// TwinCAT 3 PLC project LibraryDocumentationSample
// Title: LibraryDocumentationSample
// Company: Beckhoff Automation GmbH & Co. KG
// ProjectVersion: 1.0.0.0
// Description: This library contains various function blocks ...
// ProgramVersion: 3.1.4026.25
// project tree:
//   LibPOUs/A_Samples/ FB_DocuSample_FunctionBlock.TcPOU, FB_DocuSample_SyntaxReminder.TcPOU
//   LibPOUs/B_DocuElements/Code block/ FB_Libdoc_CodeBlock.TcPOU
//   LibPOUs/B_DocuElements/Hyperlinks/ FB_Libdoc_LinkToAnotherObject.TcPOU, FB_Libdoc_AnonymousHyperlinks.TcPOU, FB_Libdoc_Citation.TcPOU, FB_Libdoc_ExternalHyperlinks.TcPOU, FB_Libdoc_IndirectHyperlinks.TcPOU, FB_Libdoc_InlineHyperlinks.TcPOU, FB_Libdoc_InternalHyperlinks.TcPOU
//   LibPOUs/B_DocuElements/Internal Comments/ FB_Libdoc_InternalComments.TcPOU
//   LibPOUs/B_DocuElements/Font style/ FB_Libdoc_FontStyle.TcPOU
//   LibPOUs/B_DocuElements/Hyperlinks/Footnotes/ FB_Libdoc_AutomaticallyNumberedFootnotes.TcPOU, FB_Libdoc_AutomaticallySymbolFootnotes.TcPOU, FB_Libdoc_ManuallyAndAutomaticallyNumberedFootnotes.TcPOU, FB_Libdoc_ManuallyNumberedFootnotes.TcPOU, FB_Libdoc_NamedAutomaticallyNumberedFootnotes.TcPOU
//   LibPOUs/B_DocuElements/Images/ FB_Libdoc_Images.TcPOU
//   LibPOUs/B_DocuElements/Lists/ FB_Libdoc_DefinitionList.TcPOU, FB_Libdoc_FieldList.TcPOU, FB_Libdoc_OrderedNumberedEnumerationList.TcPOU, FB_Libdoc_UnorderedEnumerationList.TcPOU
//   LibPOUs/B_DocuElements/Note elements/ FB_Libdoc_SpecificNotes.TcPOU, FB_Libdoc_GenericNotes.TcPOU
//   LibPOUs/B_DocuElements/Comment structure/ FB_Libdoc_Sections.TcPOU, FB_Libdoc_Transitions.TcPOU
//   LibPOUs/B_DocuElements/Substitution/ FB_Libdoc_Substitution_ReplacementText.TcPOU, FB_Libdoc_Substitution_Images.TcPOU
//   LibPOUs/B_DocuElements/Tables/ FB_Libdoc_CSVTable.TcPOU, FB_Libdoc_GridTable.TcPOU, FB_Libdoc_ListTable.TcPOU, FB_Libdoc_SimpleTables.TcPOU
//   LibPOUs/B_DocuElements/Text blocks/ FB_Libdoc_LineBlock.TcPOU, FB_Libdoc_Paragraph.TcPOU, FB_Libdoc_BlockQuote.TcPOU

// ---- LibPOUs/A_Samples/FB_DocuSample_FunctionBlock.TcPOU
(* 
:Description: This function block represents <...> and can be used for <...> ...
:Instructions for use: How to use this FB ...

Version history:

+-------------+------------+----------------+----------+------------------------------------------+
|Date         | Version    | created under  | Author   | Remark                                   |
+=============+============+================+==========+==========================================+
|2017-07-04   | 1.0.0.0    | V3.1.4022.0    | S.H.     | Performance optimization                 |
+-------------+------------+----------------+----------+------------------------------------------+
|2019-01-11   | 1.1.0.0    | V3.1.4022.27   | K.F.     | Bug fix: Output calculation corrected    |
+-------------+------------+----------------+----------+------------------------------------------+
*)

FUNCTION_BLOCK FB_DocuSample_FunctionBlock
VAR_INPUT
    nVarInA : INT;       //First input variable
    nVarInB : INT := 5;  //Second input variable
END_VAR
VAR_OUTPUT
    nVarOut : INT;       //Output variable
END_VAR

END_FUNCTION_BLOCK

// ---- LibPOUs/A_Samples/FB_DocuSample_SyntaxReminder.TcPOU
(*
=================================================
The reStructuredText Cheat Sheet: Syntax Reminder
=================================================
:Info: See <https://infosys.beckhoff.de/.
:Author: Beckhoff <support@beckhoff.com>
:Date: 2017-12-14

.. NOTE:: This syntax reminder is based on the docutils documentation

Section Structure
=================

A reStructuredText comment is made up of body elements, and may be
structured into sections. Section titles are underlined or overlined and underlined.
Sections contain body elements and/or subsections.

Paragraphs are flush-left and separated by blank lines.

Body Elements
=============
Grid table:

+--------------------------------+-------------------------------------+
|Block quotes consist of         |Literal block, preceded by "::"::    |
|indented body elements:         |                                     |
|                                |    If (a=TRUE) Then                 |
|    Block quotes are indented.  |      b=3                            |
|                                |                                     |
+--------------------------------+-------------------------------------+
|| Line blocks preserve line breaks and indents.                       |
||    Useful for adornment-free lists;                                 |
||    long lines can be wrapped                                        |
|     with continuation lines.                                         |
+----------------------------------------------------------------------+

Simple table:

================  ========================================================
List Type         Examples
================  ========================================================
Bullet list       - This is a bullet list
                  - Items begin with "-", "+", or "*"
Enumerated list   1. This is an enumerated list.
                  2. Items use any variation of "1.", "A)", and "(i)"
                  #. Item can also be auto-enumerated
Definition list   Term is flush-left : optional classifier
                      Definition is indented, no blank line between
                      continue
Field list        :Field name: field body
================  ========================================================

Inline Markup
=============
*emphasis*, **strong emphasis**, ``inline literal text``

| Standalone hyperlink: http://beckhoff.de
| Named reference: Beckhoff_
| Anonymous reference: `Anonymous reference`__
| Footnote reference: [1]_
| Citation reference: [CIT2002]_
| Substitution: |substitution|
| Inline internal target: `Inline internal target`_

Explicit Markup
================

================  ========================================================
Explicit Markup       Examples (visible in the source code)
================  ========================================================
Footnote          .. [1] Manually numbered or [#] auto-numbered
                        (even [#label]) or [*] auto-symbol
Citation          .. [CIT2002] This is a citation.
Hyperlink Target  .. _Beckhoff: http://beckhoff.de
                  .. _indirect target: Beckhoff_
                  .. _internal target:
Anonymous Target  __ http://beckhoff.de
Directive ("::")  .. image::, .. code::
Substitution Def  .. |substitution| replace:: This is a substitution
Comment           .. This text will not be shown
================  ========================================================

Directives
===========

================  ========================================================
Directive Name    Description
================  ========================================================
attention         Specific admonition ("caution", "danger",
                  "error", "hint", "important", "note", "tip", "warning")
admonition        Generic titled admonition
image             .. image:: C:\Tc3LibDocImages\BeckhoffLogo.png
                     :width: 40
code              .. code::

                     if(a=true) then b=3;
list-table        Create a table from a uniform two-level bullet list
csv-table         Create a table from CSV data
================  ========================================================*)

FUNCTION_BLOCK FB_DocuSample_SyntaxReminder
VAR_INPUT
    nVarInA : INT;       //First input variable
    nVarInB : INT := 5;  //Second input variable
END_VAR
VAR_OUTPUT
    nVarOut : INT;       //Output variable
END_VAR

END_FUNCTION_BLOCK

// ---- LibPOUs/B_DocuElements/Code block/FB_Libdoc_CodeBlock.TcPOU
(*

**Code block with color-coded syntax**

.. code:: 
    
    // Attempts to return the value of a boolean property.
   
    FUNCTION GetBooleanProperty : BOOL
    VAR_INPUT
        sKey: STRING;
    END_VAR

    // This structure defines a special profile.

    TYPE ST_Profile :
    STRUCT
        nId     : INT := -1;
        sBuffer : STRING(255) := 'Hello';
    END_STRUCT
    END_TYPE

**Code block with line numbering**

.. code:: 
   :number-lines: 1
    
    // Attempts to return the value of a boolean property.
   
    FUNCTION GetBooleanProperty : BOOL
    VAR_INPUT
        sKey: STRING;
    END_VAR

    // This structure defines a special profile.

    TYPE ST_Profile :
    STRUCT
        nId     : INT := -1;
        sBuffer : STRING(255) := 'Hello';
    END_STRUCT
    END_TYPE

*)

FUNCTION_BLOCK FB_Libdoc_CodeBlock
VAR_INPUT
    nVarA : INT;
    nVarB : INT;
END_VAR
VAR_OUTPUT
    nSum : INT;
END_VAR
VAR
END_VAR

END_FUNCTION_BLOCK

// ---- LibPOUs/B_DocuElements/Hyperlinks/FB_Libdoc_LinkToAnotherObject.TcPOU
(*
| It is also possible to create a reference to the documentation of another object which is also part of this library.
| For example, by clicking on this link :ref:`FB_Libdoc_InlineHyperlinks`, the documentation of this FB will be shown.
| Or you can also create a link to :ref:`FB_Libdoc_CodeBlock` which is part of another folder.

*)

FUNCTION_BLOCK FB_Libdoc_LinkToAnotherObject
VAR_INPUT
    nVarA : INT;
    nVarB : INT;
END_VAR
VAR_OUTPUT
    nSum : INT;
END_VAR
VAR
END_VAR

END_FUNCTION_BLOCK

// ---- LibPOUs/B_DocuElements/Internal Comments/FB_Libdoc_InternalComments.TcPOU
(*
This is the first paragraph.

.. Comments begin with two dots and one space. Anything can
   follow, except for the syntax of footnotes/citations,
   hyperlink targets, directives, or substitution definitions.

Since comments are not shown, this paragraph follows the previous paragraph directly.
*)

FUNCTION_BLOCK FB_Libdoc_InternalComments
VAR_INPUT
    nVarA : INT;
    nVarB : INT;
END_VAR
VAR_OUTPUT
    nSum : INT;
END_VAR
VAR
END_VAR

END_FUNCTION_BLOCK

// ---- LibPOUs/B_DocuElements/Font style/FB_Libdoc_FontStyle.TcPOU
(*
This is *emphasized text*.

This is **strong text**.

This text is an example of ``inline literals``.
*)

FUNCTION_BLOCK FB_Libdoc_FontStyle
VAR_INPUT
    nVarA : INT;
    nVarB : INT;
END_VAR
VAR_OUTPUT
    nSum : INT;
END_VAR
VAR
END_VAR

END_FUNCTION_BLOCK

// ---- LibPOUs/B_DocuElements/Hyperlinks/FB_Libdoc_AnonymousHyperlinks.TcPOU
(*
See the `Beckhoff Online Information System`__ or the `Beckhoff home page`__.

.. __: http://infosys.beckhoff.de/

.. __: http://beckhoff.de/
*)

FUNCTION_BLOCK FB_Libdoc_AnonymousHyperlinks
VAR_INPUT
    nVarA : INT;
    nVarB : INT;
END_VAR
VAR_OUTPUT
    nSum : INT;
END_VAR
VAR
END_VAR

END_FUNCTION_BLOCK

// ---- LibPOUs/B_DocuElements/Hyperlinks/FB_Libdoc_Citation.TcPOU
(*
Citation references, like [CIT2002]_. Note that citations may get rearranged, e.g., to the bottom of the "page". 

| Some sample text to get some text in between.
| Some sample text to get some text in between.
| Some sample text to get some text in between.
| Some sample text to get some text in between.
| Some sample text to get some text in between.
| Some sample text to get some text in between.

.. [CIT2002] This is the citation.  It's just like a footnote,
   except the label is textual. 

Given a citation like [this]_, one can also refer to it like this_. 

| Some sample text to get some text in between.
| Some sample text to get some text in between.
| Some sample text to get some text in between.
| Some sample text to get some text in between.
| Some sample text to get some text in between.
| Some sample text to get some text in between.

.. [this] here.

| Some sample text to get some text in between.
| Some sample text to get some text in between.
| Some sample text to get some text in between.
| Some sample text to get some text in between.
| Some sample text to get some text in between.
| Some sample text to get some text in between.

*)

FUNCTION_BLOCK FB_Libdoc_Citation
VAR_INPUT
    nVarA : INT;
    nVarB : INT;
END_VAR
VAR_OUTPUT
    nSum : INT;
END_VAR
VAR
END_VAR

END_FUNCTION_BLOCK

// ---- LibPOUs/B_DocuElements/Hyperlinks/FB_Libdoc_ExternalHyperlinks.TcPOU
(*
See the Beckhoff homepage_ for more information.

Please contact the `Beckhoff Support`_ for technical assistance.

.. _homepage: http://www.beckhoff.de
.. _Beckhoff Support: support@beckhoff.com

For more information see the `PLC Lib Tc2_System`_ and `PLC Lib Tc2_Standard`_.

.. _PLC Lib Tc2_System: https://download.beckhoff.com/download/document/automation/twincat3/TwinCAT_3_PLC_Lib_Tc2_System_EN.pdf
.. _PLC Lib Tc2_Standard: https://download.beckhoff.com/download/document/automation/twincat3/TwinCAT_3_PLC_Lib__Tc2_Standard_EN.pdf

External hyperlinks, like `Beckhoff <http://www.beckhoff.de/>`_.


**Standalone hyperlinks**

See http://www.beckhoff.de for info.

Contact support@beckhoff.com


**Embedded URIs and aliases**

See the `Beckhoff homepage <http://www.beckhoff.de>`_ for info.

This `link <Beckhoff homepage_>`_ is an alias to the link above.


See the `Beckhoff homepage`_ for info.

This link_ is an alias to the link above.

.. _Beckhoff homepage: http://www.beckhoff.de
.. _link: `Beckhoff homepage`_

*)

FUNCTION_BLOCK FB_Libdoc_ExternalHyperlinks
VAR_INPUT
    nVarA : INT;
    nVarB : INT;
END_VAR
VAR_OUTPUT
    nSum : INT;
END_VAR
VAR
END_VAR

END_FUNCTION_BLOCK

// ---- LibPOUs/B_DocuElements/Hyperlinks/FB_Libdoc_IndirectHyperlinks.TcPOU
(*

**Indirect references to an internal reference target**

This hyperlink points to target one_ and indirect to target three.

.. _one: two_
.. _two: three_
.. _three:

The hyperlink targets above point to this paragraph.

**Indirect references to an external reference target**

The `Beckhoff Information System`_ is a reference source for Beckhoff_ products

.. _Beckhoff: `Beckhoff Information System`_

.. _Beckhoff Information System: https://infosys.beckhoff.de/
*)

FUNCTION_BLOCK FB_Libdoc_IndirectHyperlinks
VAR_INPUT
    nVarA : INT;
    nVarB : INT;
END_VAR
VAR_OUTPUT
    nSum : INT;
END_VAR
VAR
END_VAR

END_FUNCTION_BLOCK

// ---- LibPOUs/B_DocuElements/Hyperlinks/FB_Libdoc_InlineHyperlinks.TcPOU
(*
| This function block is based on a _`statemachine` concept which is described in the following.
| The statemachine is based on several states.
| The proceeding always begins in the first state.
| If the last state is left, the execution restarts in the first state.
| There are so many more information necessary to describe the statemachine concept in detail.
| But as this is just a sample text to show the inline hyperlinks, we want to leave out the details.
| A rough description should be enough for the sample demonstration.
| 
| Some sample text to get some text in between.
| Some sample text to get some text in between.
| Some sample text to get some text in between.
| Some sample text to get some text in between.
| Some sample text to get some text in between.
| Some sample text to get some text in between.
| 
| Furthermore, the function block is based on another concept. This is called XY.
| It is always necessary to respect the demands of this concept.
| Especially, as it is deeply interwoven with the statemachine concept.
| Therefore, you definitely need to understand the statemachine concept first.
| Afterwards, you might understand the XY concept.
| For more information about this, see the description of the `statemachine`_.
| By clicking on this link, the Library Manager will jump to the beginning of the first paragraph where the statemachine concept is described.. 

*)

FUNCTION_BLOCK FB_Libdoc_InlineHyperlinks
VAR_INPUT
    nVarA : INT;
    nVarB : INT;
END_VAR
VAR_OUTPUT
    nSum : INT;
END_VAR
VAR
END_VAR

END_FUNCTION_BLOCK

// ---- LibPOUs/B_DocuElements/Hyperlinks/FB_Libdoc_InternalHyperlinks.TcPOU
(*

**Simple internal hyperlink target**

Clicking on this internal hyperlink will take us to the target_
below.

.. _target:

**Nesting of internal hyperlink targets**

Clicking on this internal hyperlink will take us to the `third item`_ of the bullet list.

* First list item
* Second list item

  .. _third item:

* Third list item, with hyperlink target.

**Concatentation of internal hyperlink targets**

Clicking on this internal hyperlink will take us to target1_
and clicking on this internal hyperlink will take us to target2_.
Both targets point the the same paragraph.

.. _target1:
.. _target2:

The targets "target1" and "target2" are synonyms; they both
point to this paragraph.
*)

FUNCTION_BLOCK FB_Libdoc_InternalHyperlinks
VAR_INPUT
    nVarA : INT;
    nVarB : INT;
END_VAR
VAR_OUTPUT
    nSum : INT;
END_VAR
VAR
END_VAR

END_FUNCTION_BLOCK

// ---- LibPOUs/B_DocuElements/Hyperlinks/Footnotes/FB_Libdoc_AutomaticallyNumberedFootnotes.TcPOU
(*

**Autonumbered footnotes**

Autonumbered footnotes are possible, like using [#]_ and [#]_. 

--------

.. [#] This is the first one. 

.. [#] This is the second one. 
*)

FUNCTION_BLOCK FB_Libdoc_AutomaticallyNumberedFootnotes
VAR_INPUT
    nVarA : INT;
    nVarB : INT;
END_VAR
VAR_OUTPUT
    nSum : INT;
END_VAR
VAR
END_VAR

END_FUNCTION_BLOCK

// ---- LibPOUs/B_DocuElements/Hyperlinks/Footnotes/FB_Libdoc_AutomaticallySymbolFootnotes.TcPOU
(*

Here is a symbolic 
footnote reference: [*]_ footnote reference: [*]_
footnote reference: [*]_ footnote reference: [*]_
footnote reference: [*]_ footnote reference: [*]_
footnote reference: [*]_ footnote reference: [*]_
footnote reference: [*]_ footnote reference: [*]_
footnote reference: [*]_

.. [*] This is the first footnote.
.. [*] This is the second footnote.
.. [*] This is the third footnote.
.. [*] This is the fourth footnote.
.. [*] This is the fifth footnote.
.. [*] This is the sixth footnote.
.. [*] This is the seventh footnote.
.. [*] This is the eighth footnote.
.. [*] This is the ninth footnote.
.. [*] This is the tenth footnote.
.. [*] This is the eleventh footnote.
*)

FUNCTION_BLOCK FB_Libdoc_AutomaticallySymbolFootnotes
VAR_INPUT
    nVarA : INT;
    nVarB : INT;
END_VAR
VAR_OUTPUT
    nSum : INT;
END_VAR
VAR
END_VAR

END_FUNCTION_BLOCK

// ---- LibPOUs/B_DocuElements/Hyperlinks/Footnotes/FB_Libdoc_ManuallyAndAutomaticallyNumberedFootnotes.TcPOU
(*

[2]_ will be "2" (manually numbered footnote),

[3]_ will be "3" (another manually numbered footnote),

[#]_ will be "4" (anonymous auto-numbered footnote), and

[#label]_ will be "1" (labeled auto-numbered).

--------

.. [2] This footnote is labeled manually, so its number is fixed.

.. [3] This footnote is also labeled manually, so its number is also fixed.

.. [#label] This autonumber-labeled footnote will be labeled "1".
   It is the first auto-numbered footnote and no other footnote
   with label "1" exists.  The order of the footnotes is used to
   determine numbering, not the order of the footnote references!

.. [#] This footnote will be labeled "4".  It is the second
   auto-numbered footnote, but footnote labels "1", "2", "3" are already used. 
*)

FUNCTION_BLOCK FB_Libdoc_ManuallyAndAutomaticallyNumberedFootnotes
VAR_INPUT
    nVarA : INT;
    nVarB : INT;
END_VAR
VAR_OUTPUT
    nSum : INT;
END_VAR
VAR
END_VAR

END_FUNCTION_BLOCK

// ---- LibPOUs/B_DocuElements/Hyperlinks/Footnotes/FB_Libdoc_ManuallyNumberedFootnotes.TcPOU
(*

**Numerical footnote**

Footnote references, like [5]_. Note that footnotes may get rearranged, e.g., to the bottom of the "page".

--------

.. [5] A numerical footnote. Note there's no colon after the ``]``.
*)

FUNCTION_BLOCK FB_Libdoc_ManuallyNumberedFootnotes
VAR_INPUT
    nVarA : INT;
    nVarB : INT;
END_VAR
VAR_OUTPUT
    nSum : INT;
END_VAR
VAR
END_VAR

END_FUNCTION_BLOCK

// ---- LibPOUs/B_DocuElements/Hyperlinks/Footnotes/FB_Libdoc_NamedAutomaticallyNumberedFootnotes.TcPOU
(*

**Autonumbered labeled footnotes**

They may be assigned 'autonumber labels' - for instance, [#first]_ and [#second]_. 

--------

.. [#first] a.k.a. first_ 

.. [#second] a.k.a. second_
*)

FUNCTION_BLOCK FB_Libdoc_NamedAutomaticallyNumberedFootnotes
VAR_INPUT
    nVarA : INT;
    nVarB : INT;
END_VAR
VAR_OUTPUT
    nSum : INT;
END_VAR
VAR
END_VAR

END_FUNCTION_BLOCK

// ---- LibPOUs/B_DocuElements/Images/FB_Libdoc_Images.TcPOU
(*

**Absolute or relative file path as directive argument**

Absolute path

.. image:: C:\Tc3LibDocImages\tulpis.jpg
   :width: 70px

Relative path

.. image:: ../../LibPics/penguins.jpg
   :width: 70px

**Left aligned image**

.. image:: ../../LibPics/desert.jpg
   :width: 20%

Description of the function block. Description of the function block. Description of the function block.
Description of the function block. Description of the function block. Description of the function block.
Description of the function block. Description of the function block. Description of the function block.
Description of the function block. Description of the function block. Description of the function block.

**Floating image, left aligned**

.. image:: ../../LibPics/desert.jpg
   :width: 20%
   :align: left

Description of the function block. Description of the function block. Description of the function block.
Description of the function block. Description of the function block. Description of the function block.
Description of the function block. Description of the function block. Description of the function block.
Description of the function block. Description of the function block. Description of the function block.

|
|
|
|
|

**Floating image, right aligned**

.. image:: ../../LibPics/desert.jpg
   :width: 20%
   :align: right

Description of the function block. Description of the function block. Description of the function block.
Description of the function block. Description of the function block. Description of the function block.
Description of the function block. Description of the function block. Description of the function block.
Description of the function block. Description of the function block. Description of the function block.

*)

FUNCTION_BLOCK FB_Libdoc_Images
VAR_INPUT
    nVarA : INT;
    nVarB : INT;
END_VAR
VAR_OUTPUT
    nSum : INT;
END_VAR
VAR
END_VAR

END_FUNCTION_BLOCK

// ---- LibPOUs/B_DocuElements/Lists/FB_Libdoc_DefinitionList.TcPOU
(*
Term 1
    Definition 1.

Term 2
    Definition 2, paragraph 1.

    Definition 2, paragraph 2.

Term 3 : classifier
    Definition 3.

Term 4 : classifier one : classifier two
    - Item 1
    - Item 2
*)

FUNCTION_BLOCK FB_Libdoc_DefinitionList
VAR_INPUT
    nVarA : INT;
    nVarB : INT;
END_VAR
VAR_OUTPUT
    nSum : INT;
END_VAR
VAR
END_VAR

END_FUNCTION_BLOCK

// ---- LibPOUs/B_DocuElements/Lists/FB_Libdoc_FieldList.TcPOU
(*
:Organization: Beckhoff Automation GmbH & Co. KG
:Contact: info@beckhoff.de
:Address: | Hülshorstweg 20
          | 33415 Verl
          | Germany
:Authors: - Me
          - Myself
          - I
:Version: 1.0
:Status: released
:Date: 2017-12-07

:Copyright:
 © Beckhoff Automation GmbH & Co. KG, Germany.
 The reproduction, distribution and utilization of this document as well as 
 the communication of its contents to others without express authorization are prohibited.
 Offenders will be held liable for the payment of damages. 
 All rights reserved in the event of the grant of a patent, utility model or design.
:Abstract: topic
:Indentation:
 Since the field marker may be quite long, the second
 and subsequent lines of the field body do not have to line up
 with the first line, but they must be indented relative to the
 field name marker, and they must line up with each other.
:LongLongFieldname: Since the field marker is quite long,
                    the field body is shown in the line after the marker.
:Parameter nIn: Integer
:Parameter nVarB: Integer
:*Parameter nVarC*: Integer
:``Parameter nVarD``: Integer
*)

FUNCTION_BLOCK FB_Libdoc_FieldList
VAR_INPUT
    nVarA : INT;
    nVarB : INT;
END_VAR
VAR_OUTPUT
    nSum : INT;
END_VAR
VAR
END_VAR

END_FUNCTION_BLOCK

// ---- LibPOUs/B_DocuElements/Lists/FB_Libdoc_OrderedNumberedEnumerationList.TcPOU
(*
1) This is the first item in the list.

   (a) This is the first subitem (1a).
   (b) This is the second subitem (1b).

2) This is the second item in the list.

   (a) This is the first subitem (2a).
   (b) This is the second subitem (2b).

#) This item is auto-enumerated.
*)

FUNCTION_BLOCK FB_Libdoc_OrderedNumberedEnumerationList
VAR_INPUT
    nVarA : INT;
    nVarB : INT;
END_VAR
VAR_OUTPUT
    nSum : INT;
END_VAR
VAR
END_VAR

END_FUNCTION_BLOCK

// ---- LibPOUs/B_DocuElements/Lists/FB_Libdoc_UnorderedEnumerationList.TcPOU
(*
This paragraph is not part of the list.

- This is the first bullet list item.  The blank line above the
  first list item is required; blank lines between list items
  (such as below this paragraph) are optional.

  - This is a sublist. The bullet lines up with the left edge
    of the text blocks above. A sublist is a new list so
    requires a blank line above. A blank line below is optional.

  - This is a sublist. The bullet lines up with the left edge
    of the text blocks above. A sublist is a new list so
    requires a blank line above. A blank line below is optional.

- This is the second item of the main list.

- This is the third item of the main list.

This paragraph is not part of the list.
*)

FUNCTION_BLOCK FB_Libdoc_UnorderedEnumerationList
VAR_INPUT
    nVarA : INT;
    nVarB : INT;
END_VAR
VAR_OUTPUT
    nSum : INT;
END_VAR
VAR
END_VAR

END_FUNCTION_BLOCK

// ---- LibPOUs/B_DocuElements/Note elements/FB_Libdoc_SpecificNotes.TcPOU
(*
.. note:: This is a note admonition.
   This is the second line of the first paragraph.

   - The note contains all indented body elements
     following.
   - It includes this bullet list.
*)

FUNCTION_BLOCK FB_Libdoc_SpecificNotes
VAR_INPUT
    nVarA : INT;
    nVarB : INT;
END_VAR
VAR_OUTPUT
    nSum : INT;
END_VAR
VAR
END_VAR

END_FUNCTION_BLOCK

// ---- LibPOUs/B_DocuElements/Note elements/FB_Libdoc_GenericNotes.TcPOU
(*
.. admonition:: And, by the way...

   You can make up your own admonition too.
*)

FUNCTION_BLOCK FB_Libdoc_GenericNotes
VAR_INPUT
    nVarA : INT;
    nVarB : INT;
END_VAR
VAR_OUTPUT
    nSum : INT;
END_VAR
VAR
END_VAR

END_FUNCTION_BLOCK

// ---- LibPOUs/B_DocuElements/Comment structure/FB_Libdoc_Sections.TcPOU
(*
Section Title
-------------
This document consists of two main sections and several subsections. All text blocks up to the next title of the same or higher level
are included in a section (or subsection, etc.).

================
1. Section Title
================
Sections are identified through their titles, which are marked up with adornment:
"underlines" below the title text, or underlines and matching "overlines" above the title.

-----------------
1.1 Section Title
-----------------
A document must be consistent in its use of section titles: once a hierarchy of title styles is established,
sections must use that hierarchy.
Rather than imposing a fixed number and order of section title adornment styles,
the order enforced will be the order as encountered.
The first style encountered will be an outermost title, the second style will be a subtitle,
the third will be a subsubtitle, and so on.

1.2.1 Section Title
===================
Underline-only adornment styles are distinct
from overline-and-underline styles that use the same character. 

1.2.1.1 Section Title
*********************
An underline/overline is a single repeated punctuation character that begins in column 1
and forms a line extending at least as far as the right edge of the title text.

1.2.1.2 Section Title
*********************

1.2.2 Section Title
===================

-----------------
1.2 Section Title
-----------------

=================
2. Section Title
=================

-----------------
2.1 Section Title
-----------------
*)

FUNCTION_BLOCK FB_Libdoc_Sections
VAR_INPUT
    nVarA : INT;
    nVarB : INT;
END_VAR
VAR_OUTPUT
    nSum : INT;
END_VAR
VAR
END_VAR

END_FUNCTION_BLOCK

// ---- LibPOUs/B_DocuElements/Comment structure/FB_Libdoc_Transitions.TcPOU
(*
A transition marker is a horizontal line 
of 4 or more repeated punctuation characters. 

------------ 

A transition should not begin or end a section or document,
nor should two transitions be immediately adjacent.
*)

FUNCTION_BLOCK FB_Libdoc_Transitions
VAR_INPUT
    nVarA : INT;
    nVarB : INT;
END_VAR
VAR_OUTPUT
    nSum : INT;
END_VAR
VAR
END_VAR

END_FUNCTION_BLOCK

// ---- LibPOUs/B_DocuElements/Substitution/FB_Libdoc_Substitution_ReplacementText.TcPOU
(*
**Substitution in paragraphs**

|RST|_ is an easy-to-read, what-you-see-is-what-you-get plaintext markup syntax.
Among others it is useful for library documentation. If the |RST| option is activated,
comments written in |RST| will be shown in the Documentation tab of the library manager in an attractive format.
|RST| is a little annoying to type over and over and spelling out the
bicapitalized word |RST| every time isn't really necessary for |RST| source readability.

.. |RST| replace:: reStructuredText
.. _RST: https://infosys.beckhoff.de/


This is a simple |substitution reference|. It will be replaced by
the processing system.

This is a |substitution and hyperlink reference|_. In
addition to being replaced, the replacement text or element will
refer to the "substitution and hyperlink reference" target.

.. |substitution reference| replace:: example of substitution 
.. |substitution and hyperlink reference| replace:: combination of substitution and hyperlink reference
.. _substitution and hyperlink reference: https://beckhoff.de/
*)

FUNCTION_BLOCK FB_Libdoc_Substitution_ReplacementText
VAR_INPUT
    nVarA : INT;
    nVarB : INT;
END_VAR
VAR_OUTPUT
    nSum : INT;
END_VAR
VAR
END_VAR

END_FUNCTION_BLOCK

// ---- LibPOUs/B_DocuElements/Substitution/FB_Libdoc_Substitution_Images.TcPOU
(*
**Substitution in paragraphs**

Images are a common use for substitution references: |Beckhoff|_.

.. |Beckhoff| image:: ../../LibPics/BeckhoffLogo.png
 :height: 16
 :width: 64
.. _Beckhoff: http://www.beckhoff.de/

The |safety| symbol indicates a hazardous situation which,
if not avoided, could result in minor or moderate injury.

.. |safety| image:: ../../LibPics/safetysymbol.png


**Substitution in lists or tables**

* |Run mode| Run mode
* |Stop mode| Stop mode
* |Config mode| Config mode

============= ======
Symbol        Status
============= ======
|Run mode|    Run mode
|Stop mode|   Stop mode
|Config mode| Config mode
============= ======

.. |Run mode| image:: ../../LibPics/tc3runmode.png
.. |Stop mode| image:: ../../LibPics/tc3stopmode.png
.. |Config mode| image:: ../../LibPics/tc3configmode.png
*)

FUNCTION_BLOCK FB_Libdoc_Substitution_Images
VAR_INPUT
    nVarA : INT;
    nVarB : INT;
END_VAR
VAR_OUTPUT
    nSum : INT;
END_VAR
VAR
END_VAR

END_FUNCTION_BLOCK

// ---- LibPOUs/B_DocuElements/Tables/FB_Libdoc_CSVTable.TcPOU
(*
.. csv-table:: Property list
   :header: "Items", "Property 1", "Property 2", "Property 3"
   :widths: 10, 15, 15, 15

   "Item 1", 1.67, angular, red
   "Item 2", "not specified", round, blue

|

.. csv-table:: Property list
   :header-rows: 1
   :widths: 10, 15, 15, 15

   "Items", "Property 1", "Property 2", "Property 3"
   "Item 1", 1.67, angular, red
   "Item 2", "not specified", round, blue
*)

FUNCTION_BLOCK FB_Libdoc_CSVTable
VAR_INPUT
    nVarA : INT;
    nVarB : INT;
END_VAR
VAR_OUTPUT
    nSum : INT;
END_VAR
VAR
END_VAR

END_FUNCTION_BLOCK

// ---- LibPOUs/B_DocuElements/Tables/FB_Libdoc_GridTable.TcPOU
(*
+------------------------+------------+----------+----------+
| Header row, column 1   | Header 2   | Header 3 | Header 4 |
| (header rows optional) |            |          |          |
+========================+============+==========+==========+
| body row 1, column 1   | column 2   | column 3 | column 4 |
+------------------------+------------+----------+----------+
| body row 2             | Cells may span columns.          |
+------------------------+------------+---------------------+
| body row 3             | Cells may  | - Table cells       |
+------------------------+ span rows. | - contain           |
| body row 4             |            | - body elements.    |
+------------------------+------------+---------------------+
*)

FUNCTION_BLOCK FB_Libdoc_GridTable
VAR_INPUT
    nVarA : INT;
    nVarB : INT;
END_VAR
VAR_OUTPUT
    nSum : INT;
END_VAR
VAR
END_VAR

END_FUNCTION_BLOCK

// ---- LibPOUs/B_DocuElements/Tables/FB_Libdoc_ListTable.TcPOU
(*
.. list-table:: Property list
    :widths: 50 50 50
    :header-rows: 1

    * - Items
      - Property 1
      - Property 2
    * - Item 1
      - angular
      - red
    * - Item 2
      - round
      - blue
*)

FUNCTION_BLOCK FB_Libdoc_ListTable
VAR_INPUT
    nVarA : INT;
    nVarB : INT;
END_VAR
VAR_OUTPUT
    nSum : INT;
END_VAR
VAR
END_VAR

END_FUNCTION_BLOCK

// ---- LibPOUs/B_DocuElements/Tables/FB_Libdoc_SimpleTables.TcPOU
(*
=====  =====  =======
  A      B    A and B
=====  =====  =======
False  False  False
True   False  False
False  True   False
True   True   True
=====  =====  =======

|

=====  =====  ======
   Inputs     Output
------------  ------
  A      B    A or B
=====  =====  ======
False  False  False
True   False  True
False  True   True
True   True   True
=====  =====  ======

|

=====  =====  ======
   Inputs     Output
------------  ------
  A      B    A or B
=====  =====  ======
False  False  False
       False  True
False  True   True
True   True   True
=====  =====  ======

|

=====  =====
Col 1  Col 2
=====  =====
1      Second column of row 1.
2      Second column of row 2.
       Second line of paragraph.
3      Second column of row 2.
                             
       Second line of paragraph
4      - Second column of row 3.

       - Second item in bullet
         list (row 4, column 2).
\      Row 5; column 1 will be empty.
=====  =====
*)

FUNCTION_BLOCK FB_Libdoc_SimpleTables
VAR_INPUT
    nVarA : INT;
    nVarB : INT;
END_VAR
VAR_OUTPUT
    nSum : INT;
END_VAR
VAR
END_VAR

END_FUNCTION_BLOCK

// ---- LibPOUs/B_DocuElements/Text blocks/FB_Libdoc_LineBlock.TcPOU
(*
Line blocks are useful where the structure of lines is significant.

| Each new line begins with 
| a vertical bar ("|"). 
|     Line breaks and initial indents 
|     are preserved. 
| Continuation lines are wrapped 
  portions of long lines; they begin 
  with spaces in place of vertical bars.

    | Each new line begins with 
    | a vertical bar ("|"). 
    |     Line breaks and initial indents 
    |     are preserved. 
    | Continuation lines are wrapped 
      portions of long lines; they begin 
      with spaces in place of vertical bars.
*)

FUNCTION_BLOCK FB_Libdoc_LineBlock
VAR_INPUT
    nVarA : INT;
    nVarB : INT;
END_VAR
VAR_OUTPUT
    nSum : INT;
END_VAR
VAR
END_VAR

END_FUNCTION_BLOCK

// ---- LibPOUs/B_DocuElements/Text blocks/FB_Libdoc_Paragraph.TcPOU
(*
This is a paragraph.

Paragraphs line up at their left edges, and are normally separated 
by blank lines.
*)

FUNCTION_BLOCK FB_Libdoc_Paragraph
VAR_INPUT
    nVarA : INT;
    nVarB : INT;
END_VAR
VAR_OUTPUT
    nSum : INT;
END_VAR
VAR
END_VAR

END_FUNCTION_BLOCK

// ---- LibPOUs/B_DocuElements/Text blocks/FB_Libdoc_BlockQuote.TcPOU
(*
This is a top-level paragraph.

    This paragraph belongs to a first-level block quote.

    This is the second paragraph of the first-level block quote.

        This paragraph belongs to a second-level block quote.

Another top-level paragraph.

        This paragraph belongs to a second-level block quote.

    This paragraph belongs to a first-level block quote. The
    second-level block quote above is inside this first-level
    block quote.
*)

FUNCTION_BLOCK FB_Libdoc_BlockQuote
VAR_INPUT
    nVarA : INT;
    nVarB : INT;
END_VAR
VAR_OUTPUT
    nSum : INT;
END_VAR
VAR
END_VAR

END_FUNCTION_BLOCK
